(* PLC project Unnamed, Unknown Unnamed 1 *)
(* stored: creationDateTime 2026-08-31T18:43:54, modificationDateTime 2026-08-31T18:43:54 *)

FUNCTION_BLOCK TON
  VAR_OUTPUT
    Q : BOOL;
    ET : TIME;
  END_VAR
  VAR_INPUT
    IN : BOOL;
    PT : TIME;
  END_VAR

END_FUNCTION_BLOCK

PROGRAM main
  VAR
    stop : BOOL;
    start : BOOL;
    motor_run : BOOL;
    star : BOOL;
    TON0 : TON;
    delta : BOOL;
    TON1 : TON;
    overload : BOOL;
    red_lamp : BOOL;
  END_VAR

(* LD diagram, written out as Structured Text *)
motor_run := NOT stop AND NOT overload AND (start OR motor_run);
star := motor_run AND NOT TON0.Q AND NOT overload;
delta := motor_run AND TON1.Q AND NOT star AND NOT overload;
red_lamp := overload;
TON0(IN := motor_run, PT := T#5s);
TON1(IN := TON0.Q, PT := T#500ms);
END_PROGRAM

CONFIGURATION Config0
  RESOURCE Res0 ON PLC
    TASK task0(INTERVAL := T#20ms, PRIORITY := 1);
    PROGRAM instance0 WITH task0 : main;
  END_RESOURCE
END_CONFIGURATION
